// Compteurs de maintenance persistants d'un élément de pool (docs/11 § 5, D92) et leur restauration (docs/02 § 7.4)
INTERFACE I_Maintained

// Objet du projet auquel appartiennent les compteurs (persistant : survit au redémarrage du PLC)
PROPERTY StableId : UDINT
GET
END_GET
END_PROPERTY

PROPERTY ActionCount : UDINT
GET
END_GET
END_PROPERTY

PROPERTY ErrorCount : UDINT
GET
END_GET
END_PROPERTY

PROPERTY MotionHours : LREAL
GET
END_GET
END_PROPERTY

METHOD RestoreCounters
VAR_INPUT
    nActions : UDINT;
    nErrors : UDINT;
    fHours : LREAL;
END_VAR
END_METHOD

END_INTERFACE

(* stored: Version 1.1.0.1, ProductVersion 3.1.4024.12
   Itf I_Maintained: Id {248e718f-e62e-564a-8032-8cf03bdfb463}
   Property StableId: Id {35146746-a7c7-551b-ad2d-3564b28cae99}
   Get Get: Id {68fe4d34-5c05-59e3-a9d1-63eedaaa1943}
   Property ActionCount: Id {04ab5a85-b0dd-541d-b5d4-ad7727089020}
   Get Get: Id {b5ba7830-15dd-5790-8a84-517dbf228a5f}
   Property ErrorCount: Id {6d0e1e1c-95fd-56b9-8586-f4cff2c828c2}
   Get Get: Id {bf9115bd-d6bc-5d9e-928b-4d0cbb760a20}
   Property MotionHours: Id {67f133e4-ba07-52fb-84ce-c04e6075becf}
   Get Get: Id {69cd8233-8b60-5b40-beb4-1a0b9050ccad}
   Method RestoreCounters: Id {f94199f3-827a-524b-b63b-112bc47f5b5a} *)
